TYPE ST_Alias :
STRUCT
    {attribute 'pytmc' := '
        alias: .ATHM
        pv: bTestATHM
    '}
     bTestATHM : BOOL;

    {attribute 'pytmc' := '
        alias: .CNEN
        pv: bTestCNEN
    '}
     bTestCNEN : BOOL;
    {attribute 'pytmc' := '
        pv: nTest64LINT
        io: io
        field: DESC Start an AbsoluteMove
    '}
END_STRUCT
END_TYPE

(* stored: Version 1.1.0.1
   DUT ST_Alias: Id {3b89bffe-1d15-45a2-a122-6c44d0d9528d} *)
